FUNCTION_BLOCK FB_MotorControl
VAR_INPUT
	bEnable : BOOL;
    bForward : BOOL;
    bBackward : BOOL;
    bForwardLimit : BOOL;
    bBackwardLimit : BOOL;
END_VAR

VAR_OUTPUT
	bMotorRun : BOOL;
    bMotorDirection : BOOL;
END_VAR

VAR
	bAllowedForward : BOOL;
    bAllowedBackward : BOOL;
	bDirectionChange : BOOL;
	bDelayElapsed : BOOL;
	
	fbDirectionDelay: TON;
	tDirectionElapsed : TIME;
END_VAR

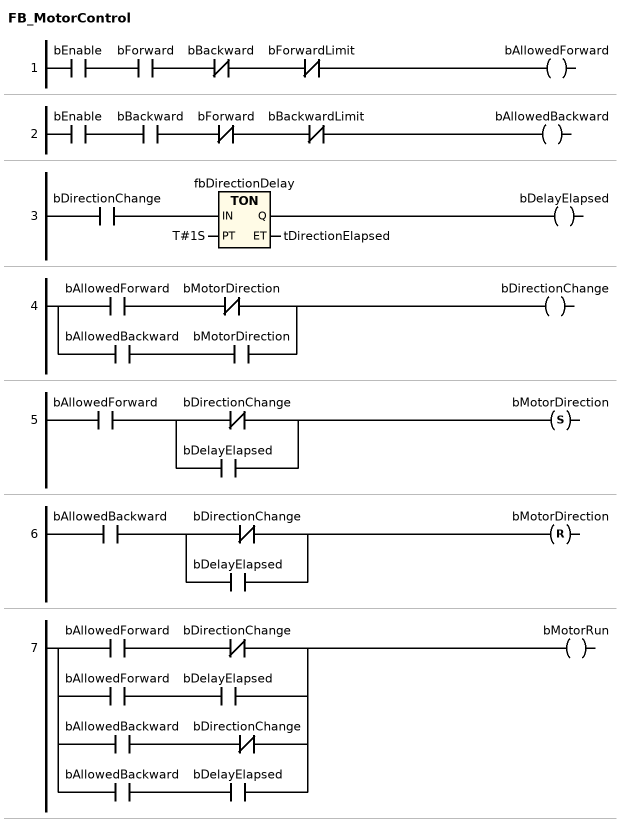
// NETWORK 1
bAllowedForward := bEnable AND bForward AND NOT bBackward AND NOT bForwardLimit;

// NETWORK 2
bAllowedBackward := bEnable AND bBackward AND NOT bForward AND NOT bBackwardLimit;

// NETWORK 3
fbDirectionDelay(IN := bDirectionChange, PT := T#1S, ET => tDirectionElapsed); // TON
bDelayElapsed := fbDirectionDelay.Q;

// NETWORK 4
bDirectionChange := bAllowedForward AND NOT bMotorDirection OR bAllowedBackward AND bMotorDirection;

// NETWORK 5
bMotorDirection S= bAllowedForward AND (NOT bDirectionChange OR bDelayElapsed);

// NETWORK 6
bMotorDirection R= bAllowedBackward AND (NOT bDirectionChange OR bDelayElapsed);

// NETWORK 7
bMotorRun := bAllowedForward AND NOT bDirectionChange OR bAllowedForward AND bDelayElapsed OR bAllowedBackward AND NOT bDirectionChange OR bAllowedBackward AND bDelayElapsed;

END_FUNCTION_BLOCK

(* stored: Version 1.1.0.1
   POU FB_MotorControl: Id {e48fc4d2-27e1-40bb-971d-9ba002d1f392}, SpecialFunc None *)
